// TIA Portal V20 export
// export: Created 2026-10-19T18:42:36.9079896Z, ExportSetting WithDefaults, DisplayName Totally Integrated Automation Portal, DisplayVersion V20 Update 6, DisplayName TIA Portal Openness, DisplayVersion V20 Update 6, DisplayName TIA Portal Version Control Interface, DisplayVersion V20 Update 6, DisplayName SINAMICS Startdrive Advanced, DisplayVersion V20 SP1, DisplayName SINAMICS Startdrive G130, G150, S120, S150, SINAMICS MV, G220, S200, S210, DisplayVersion V20 SP1, DisplayName SINAMICS Startdrive G110M, G120, G120C, G120D, G120P, G115D, DisplayVersion V20 SP1, DisplayName STEP 7 Professional, DisplayVersion V20 Update 6, DisplayName STEP 7 Safety, DisplayVersion V20 Update 2, DisplayName WinCC Basic/Comfort/Advanced, DisplayVersion V20 Update 6, DisplayName WinCC Unified, DisplayVersion V20 Update 6
FUNCTION_BLOCK "Remote_Panel"   // FB17, F_LAD
{ S7_Optimized_Access := 'TRUE' }
VERSION : 0.1
// stored: AutoNumber true, IsIECCheckEnabled false, UDAEnableTagReadback false
   VAR_INPUT
      ID : Int;
      Overtravel_Lower_limit : Bool;
      Overtravel_Upper_limit : Bool;
      Estop : Bool;
      Reset : Bool;
      Chain_Slack_1 : Bool;
      Chain_Slack_2 : Bool;
      Chain_Slack_3 : Bool;
      Chain_Slack_4 : Bool;
      "Light Guards 1" : Bool;
      "Light Guards 2" : Bool;
      Gate_1 : Bool;
      Gate_2 : Bool;
      EStop_Lock_1 : Bool;
      EStop_Lock_2 : Bool;
      Lock_Secured_1 : Bool;
      Lock_Secured_2 : Bool;
      "EStop Level 1" : Bool;
      "EStop Level 2" : Bool;
      "EStop Level 3" : Bool;
      "EStop Level 4" : Bool;
      "EStop Level 5" : Bool;
      "EStop Level 6" : Bool;
      Bypass : "F_Bypass_RemotePanel";
   END_VAR
   VAR_OUTPUT
      Safety_OK : Bool;
      Bypass_Warning : Bool;
      "STO VTD - CH1" : Bool;
      "STO VTD - CH2" : Bool;
      ACK { ExternalAccessible := 'False'; ExternalVisible := 'False'; ExternalWritable := 'False'} : Bool;
      L1_OK : Bool;
      L2_OK : Bool;
      L3_OK : Bool;
      L4_OK : Bool;
      L5_OK : Bool;
      L6_OK : Bool;
   END_VAR
   VAR
      Overtravel_Lower_Limit_DB : ESTOP1;
      Overtravel_Upper_Limit_DB : ESTOP1;
      Estop_Cabinet_DB : ESTOP1;
      Chain_Slack_1_DB : ESTOP1;
      Chain_Slack_2_DB : ESTOP1;
      Chain_Slack_3_DB : ESTOP1;
      Chain_Slack_4_DB : ESTOP1;
      "Light_Guards 1" : ESTOP1;
      "Light_Guards 2" : ESTOP1;
      Gate_1_DB : ESTOP1;
      Gate_2_DB : ESTOP1;
      EStop_Lock_1_DB : ESTOP1;
      EStop_Lock_2_DB : ESTOP1;
      Lock_Secured_1_DB : ESTOP1;
      Lock_Secured_2_DB : ESTOP1;
      "EStop Level 1_DB" : ESTOP1;
      "EStop Level 2_DB" : ESTOP1;
      "EStop Level 3_DB" : ESTOP1;
      "EStop Level 4_DB" : ESTOP1;
      "EStop Level 5_DB" : ESTOP1;
      "EStop Level 6_DB" : ESTOP1;
   END_VAR
   VAR_TEMP
      EStop_Levels_OK : Bool;
   END_VAR
BEGIN

REGION Network 1: RESET CABINET
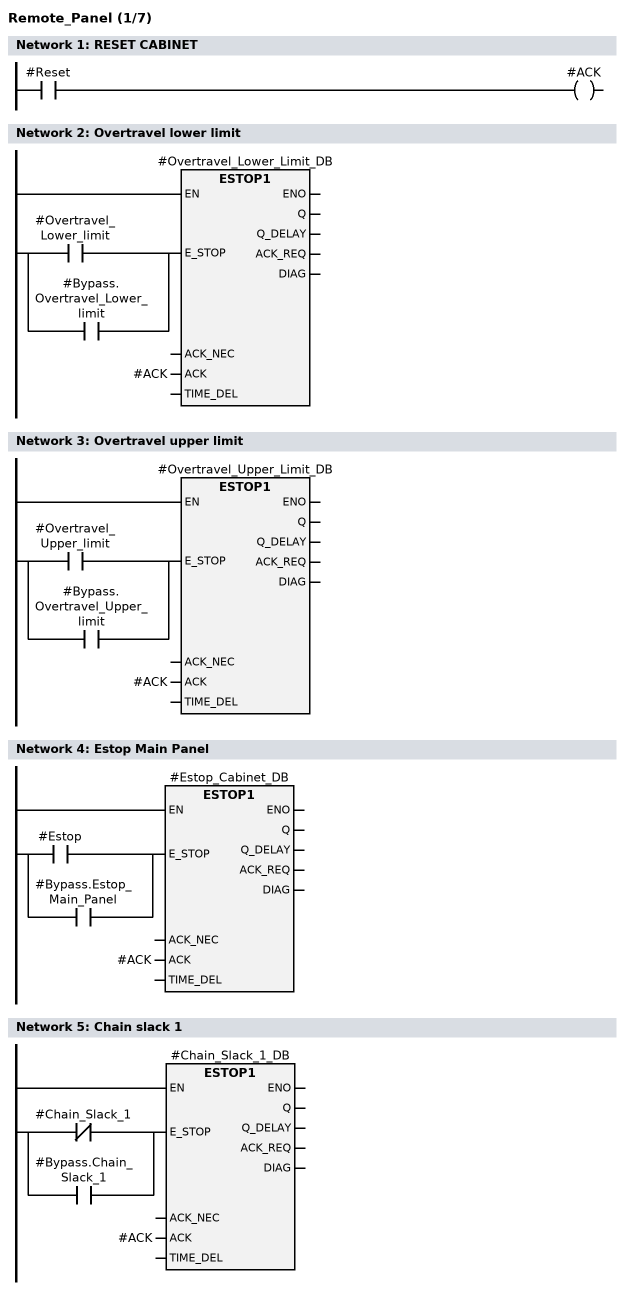
   RUNG wire#powerrail
      Contact( #Reset )
      Coil( #ACK )
   END_RUNG
   // the same network as SCL:
   #ACK := #Reset;
END_REGION

REGION Network 2: Overtravel lower limit
   RUNG wire#powerrail
      #Overtravel_Lower_Limit_DB.ESTOP1(E_STOP := wire#w1, ACK_NEC :=, ACK := #ACK, TIME_DEL :=, Q =>, Q_DELAY =>, ACK_REQ =>, DIAG =>)
   END_RUNG
   RUNG wire#powerrail
      Contact( #Overtravel_Lower_limit )
   END_RUNG wire#w1
   RUNG wire#powerrail
      Contact( #Bypass.Overtravel_Lower_limit )
   END_RUNG wire#w1
   // the same network as SCL:
   #Overtravel_Lower_Limit_DB(E_STOP := #Overtravel_Lower_limit OR #Bypass.Overtravel_Lower_limit, ACK := #ACK);   // ESTOP1
END_REGION

REGION Network 3: Overtravel upper limit
   RUNG wire#powerrail
      #Overtravel_Upper_Limit_DB.ESTOP1(E_STOP := wire#w1, ACK_NEC :=, ACK := #ACK, TIME_DEL :=, Q =>, Q_DELAY =>, ACK_REQ =>, DIAG =>)
   END_RUNG
   RUNG wire#powerrail
      Contact( #Overtravel_Upper_limit )
   END_RUNG wire#w1
   RUNG wire#powerrail
      Contact( #Bypass.Overtravel_Upper_limit )
   END_RUNG wire#w1
   // the same network as SCL:
   #Overtravel_Upper_Limit_DB(E_STOP := #Overtravel_Upper_limit OR #Bypass.Overtravel_Upper_limit, ACK := #ACK);   // ESTOP1
END_REGION

REGION Network 4: Estop Main Panel
   RUNG wire#powerrail
      #Estop_Cabinet_DB.ESTOP1(E_STOP := wire#w1, ACK_NEC :=, ACK := #ACK, TIME_DEL :=, Q =>, Q_DELAY =>, ACK_REQ =>, DIAG =>)
   END_RUNG
   RUNG wire#powerrail
      Contact( #Estop )
   END_RUNG wire#w1
   RUNG wire#powerrail
      Contact( #Bypass.Estop_Main_Panel )
   END_RUNG wire#w1
   // the same network as SCL:
   #Estop_Cabinet_DB(E_STOP := #Estop OR #Bypass.Estop_Main_Panel, ACK := #ACK);   // ESTOP1
END_REGION

REGION Network 5: Chain slack 1
   RUNG wire#powerrail
      #Chain_Slack_1_DB.ESTOP1(E_STOP := wire#w1, ACK_NEC :=, ACK := #ACK, TIME_DEL :=, Q =>, Q_DELAY =>, ACK_REQ =>, DIAG =>)
   END_RUNG
   RUNG wire#powerrail
      I_Contact( #Chain_Slack_1 )
   END_RUNG wire#w1
   RUNG wire#powerrail
      Contact( #Bypass.Chain_Slack_1 )
   END_RUNG wire#w1
   // the same network as SCL:
   #Chain_Slack_1_DB(E_STOP := NOT #Chain_Slack_1 OR #Bypass.Chain_Slack_1, ACK := #ACK);   // ESTOP1
END_REGION

REGION Network 6: Chain slack 2
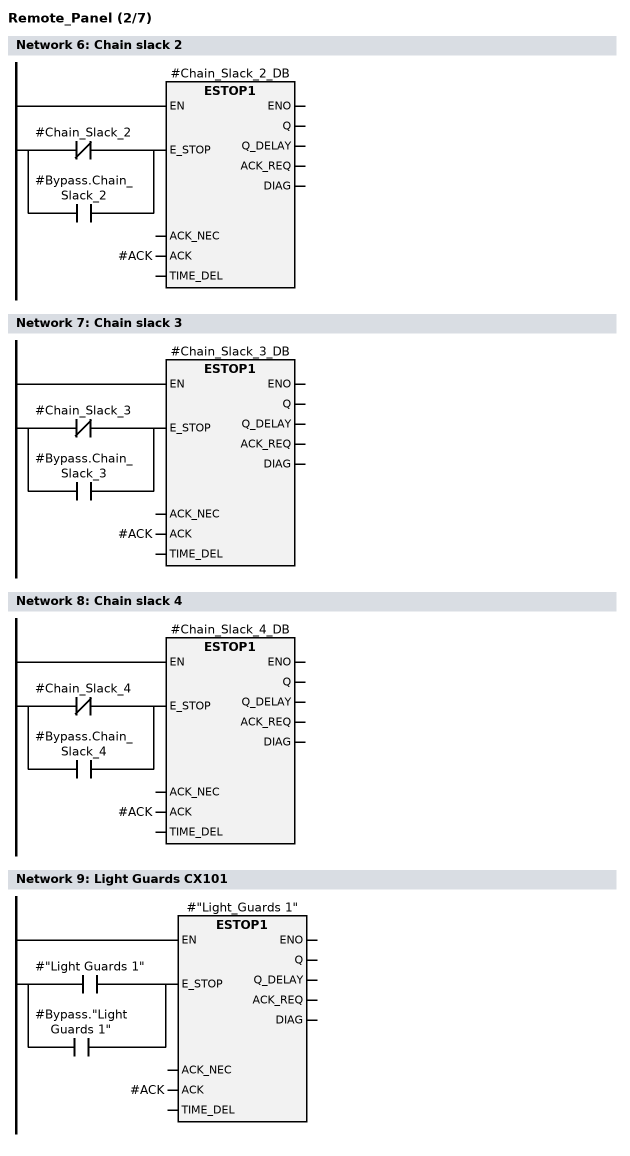
   RUNG wire#powerrail
      #Chain_Slack_2_DB.ESTOP1(E_STOP := wire#w1, ACK_NEC :=, ACK := #ACK, TIME_DEL :=, Q =>, Q_DELAY =>, ACK_REQ =>, DIAG =>)
   END_RUNG
   RUNG wire#powerrail
      I_Contact( #Chain_Slack_2 )
   END_RUNG wire#w1
   RUNG wire#powerrail
      Contact( #Bypass.Chain_Slack_2 )
   END_RUNG wire#w1
   // the same network as SCL:
   #Chain_Slack_2_DB(E_STOP := NOT #Chain_Slack_2 OR #Bypass.Chain_Slack_2, ACK := #ACK);   // ESTOP1
END_REGION

REGION Network 7: Chain slack 3
   RUNG wire#powerrail
      #Chain_Slack_3_DB.ESTOP1(E_STOP := wire#w1, ACK_NEC :=, ACK := #ACK, TIME_DEL :=, Q =>, Q_DELAY =>, ACK_REQ =>, DIAG =>)
   END_RUNG
   RUNG wire#powerrail
      I_Contact( #Chain_Slack_3 )
   END_RUNG wire#w1
   RUNG wire#powerrail
      Contact( #Bypass.Chain_Slack_3 )
   END_RUNG wire#w1
   // the same network as SCL:
   #Chain_Slack_3_DB(E_STOP := NOT #Chain_Slack_3 OR #Bypass.Chain_Slack_3, ACK := #ACK);   // ESTOP1
END_REGION

REGION Network 8: Chain slack 4
   RUNG wire#powerrail
      #Chain_Slack_4_DB.ESTOP1(E_STOP := wire#w1, ACK_NEC :=, ACK := #ACK, TIME_DEL :=, Q =>, Q_DELAY =>, ACK_REQ =>, DIAG =>)
   END_RUNG
   RUNG wire#powerrail
      I_Contact( #Chain_Slack_4 )
   END_RUNG wire#w1
   RUNG wire#powerrail
      Contact( #Bypass.Chain_Slack_4 )
   END_RUNG wire#w1
   // the same network as SCL:
   #Chain_Slack_4_DB(E_STOP := NOT #Chain_Slack_4 OR #Bypass.Chain_Slack_4, ACK := #ACK);   // ESTOP1
END_REGION

REGION Network 9: Light Guards CX101
   RUNG wire#powerrail
      #"Light_Guards 1".ESTOP1(E_STOP := wire#w1, ACK_NEC :=, ACK := #ACK, TIME_DEL :=, Q =>, Q_DELAY =>, ACK_REQ =>, DIAG =>)
   END_RUNG
   RUNG wire#powerrail
      Contact( #"Light Guards 1" )
   END_RUNG wire#w1
   RUNG wire#powerrail
      Contact( #Bypass."Light Guards 1" )
   END_RUNG wire#w1
   // the same network as SCL:
   #"Light_Guards 1"(E_STOP := #"Light Guards 1" OR #Bypass."Light Guards 1", ACK := #ACK);   // ESTOP1
END_REGION

REGION Network 10: Light Guards CX201
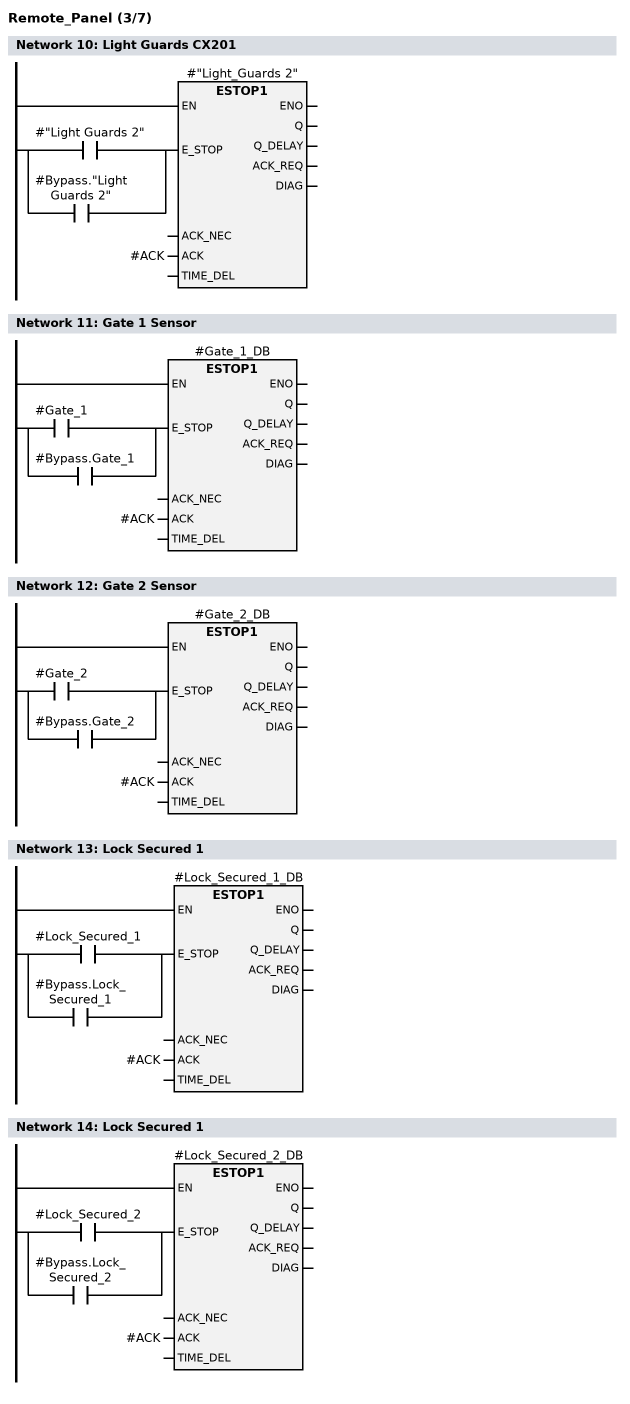
   RUNG wire#powerrail
      #"Light_Guards 2".ESTOP1(E_STOP := wire#w1, ACK_NEC :=, ACK := #ACK, TIME_DEL :=, Q =>, Q_DELAY =>, ACK_REQ =>, DIAG =>)
   END_RUNG
   RUNG wire#powerrail
      Contact( #"Light Guards 2" )
   END_RUNG wire#w1
   RUNG wire#powerrail
      Contact( #Bypass."Light Guards 2" )
   END_RUNG wire#w1
   // the same network as SCL:
   #"Light_Guards 2"(E_STOP := #"Light Guards 2" OR #Bypass."Light Guards 2", ACK := #ACK);   // ESTOP1
END_REGION

REGION Network 11: Gate 1 Sensor
   RUNG wire#powerrail
      #Gate_1_DB.ESTOP1(E_STOP := wire#w1, ACK_NEC :=, ACK := #ACK, TIME_DEL :=, Q =>, Q_DELAY =>, ACK_REQ =>, DIAG =>)
   END_RUNG
   RUNG wire#powerrail
      Contact( #Gate_1 )
   END_RUNG wire#w1
   RUNG wire#powerrail
      Contact( #Bypass.Gate_1 )
   END_RUNG wire#w1
   // the same network as SCL:
   #Gate_1_DB(E_STOP := #Gate_1 OR #Bypass.Gate_1, ACK := #ACK);   // ESTOP1
END_REGION

REGION Network 12: Gate 2 Sensor
   RUNG wire#powerrail
      #Gate_2_DB.ESTOP1(E_STOP := wire#w1, ACK_NEC :=, ACK := #ACK, TIME_DEL :=, Q =>, Q_DELAY =>, ACK_REQ =>, DIAG =>)
   END_RUNG
   RUNG wire#powerrail
      Contact( #Gate_2 )
   END_RUNG wire#w1
   RUNG wire#powerrail
      Contact( #Bypass.Gate_2 )
   END_RUNG wire#w1
   // the same network as SCL:
   #Gate_2_DB(E_STOP := #Gate_2 OR #Bypass.Gate_2, ACK := #ACK);   // ESTOP1
END_REGION

REGION Network 13: Lock Secured 1
   RUNG wire#powerrail
      #Lock_Secured_1_DB.ESTOP1(E_STOP := wire#w1, ACK_NEC :=, ACK := #ACK, TIME_DEL :=, Q =>, Q_DELAY =>, ACK_REQ =>, DIAG =>)
   END_RUNG
   RUNG wire#powerrail
      Contact( #Lock_Secured_1 )
   END_RUNG wire#w1
   RUNG wire#powerrail
      Contact( #Bypass.Lock_Secured_1 )
   END_RUNG wire#w1
   // the same network as SCL:
   #Lock_Secured_1_DB(E_STOP := #Lock_Secured_1 OR #Bypass.Lock_Secured_1, ACK := #ACK);   // ESTOP1
END_REGION

REGION Network 14: Lock Secured 1
   RUNG wire#powerrail
      #Lock_Secured_2_DB.ESTOP1(E_STOP := wire#w1, ACK_NEC :=, ACK := #ACK, TIME_DEL :=, Q =>, Q_DELAY =>, ACK_REQ =>, DIAG =>)
   END_RUNG
   RUNG wire#powerrail
      Contact( #Lock_Secured_2 )
   END_RUNG wire#w1
   RUNG wire#powerrail
      Contact( #Bypass.Lock_Secured_2 )
   END_RUNG wire#w1
   // the same network as SCL:
   #Lock_Secured_2_DB(E_STOP := #Lock_Secured_2 OR #Bypass.Lock_Secured_2, ACK := #ACK);   // ESTOP1
END_REGION

REGION Network 15: Idem Lock EStop 1
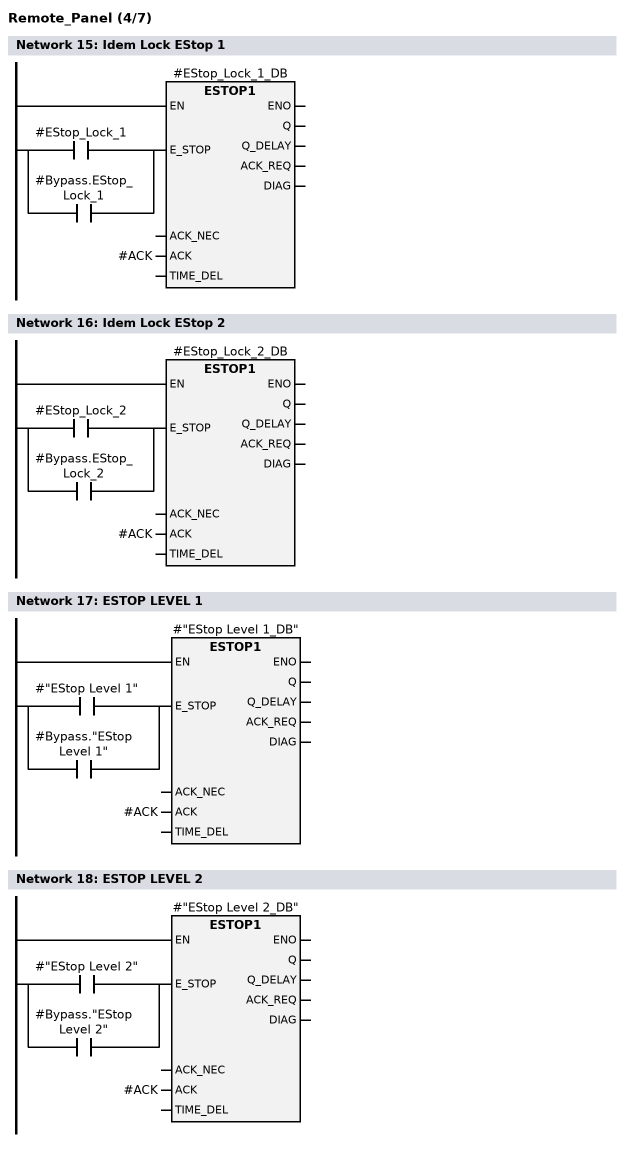
   RUNG wire#powerrail
      #EStop_Lock_1_DB.ESTOP1(E_STOP := wire#w1, ACK_NEC :=, ACK := #ACK, TIME_DEL :=, Q =>, Q_DELAY =>, ACK_REQ =>, DIAG =>)
   END_RUNG
   RUNG wire#powerrail
      Contact( #EStop_Lock_1 )
   END_RUNG wire#w1
   RUNG wire#powerrail
      Contact( #Bypass.EStop_Lock_1 )
   END_RUNG wire#w1
   // the same network as SCL:
   #EStop_Lock_1_DB(E_STOP := #EStop_Lock_1 OR #Bypass.EStop_Lock_1, ACK := #ACK);   // ESTOP1
END_REGION

REGION Network 16: Idem Lock EStop 2
   RUNG wire#powerrail
      #EStop_Lock_2_DB.ESTOP1(E_STOP := wire#w1, ACK_NEC :=, ACK := #ACK, TIME_DEL :=, Q =>, Q_DELAY =>, ACK_REQ =>, DIAG =>)
   END_RUNG
   RUNG wire#powerrail
      Contact( #EStop_Lock_2 )
   END_RUNG wire#w1
   RUNG wire#powerrail
      Contact( #Bypass.EStop_Lock_2 )
   END_RUNG wire#w1
   // the same network as SCL:
   #EStop_Lock_2_DB(E_STOP := #EStop_Lock_2 OR #Bypass.EStop_Lock_2, ACK := #ACK);   // ESTOP1
END_REGION

REGION Network 17: ESTOP LEVEL 1
   RUNG wire#powerrail
      #"EStop Level 1_DB".ESTOP1(E_STOP := wire#w1, ACK_NEC :=, ACK := #ACK, TIME_DEL :=, Q =>, Q_DELAY =>, ACK_REQ =>, DIAG =>)
   END_RUNG
   RUNG wire#powerrail
      Contact( #"EStop Level 1" )
   END_RUNG wire#w1
   RUNG wire#powerrail
      Contact( #Bypass."EStop Level 1" )
   END_RUNG wire#w1
   // the same network as SCL:
   #"EStop Level 1_DB"(E_STOP := #"EStop Level 1" OR #Bypass."EStop Level 1", ACK := #ACK);   // ESTOP1
END_REGION

REGION Network 18: ESTOP LEVEL 2
   RUNG wire#powerrail
      #"EStop Level 2_DB".ESTOP1(E_STOP := wire#w1, ACK_NEC :=, ACK := #ACK, TIME_DEL :=, Q =>, Q_DELAY =>, ACK_REQ =>, DIAG =>)
   END_RUNG
   RUNG wire#powerrail
      Contact( #"EStop Level 2" )
   END_RUNG wire#w1
   RUNG wire#powerrail
      Contact( #Bypass."EStop Level 2" )
   END_RUNG wire#w1
   // the same network as SCL:
   #"EStop Level 2_DB"(E_STOP := #"EStop Level 2" OR #Bypass."EStop Level 2", ACK := #ACK);   // ESTOP1
END_REGION

REGION Network 19: ESTOP LEVEL 3
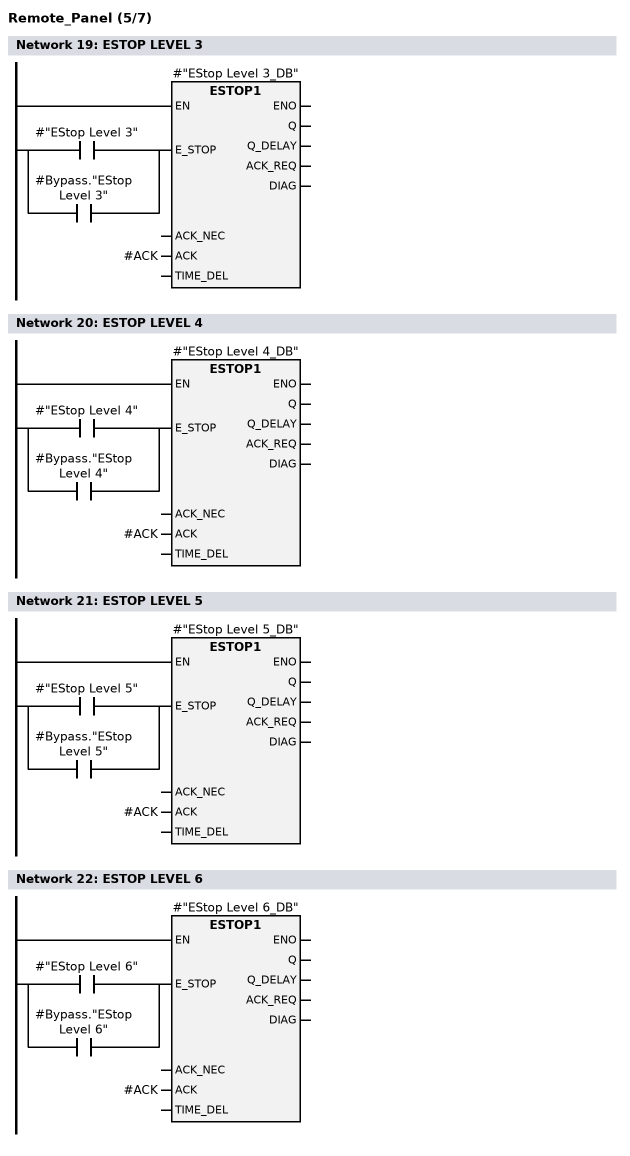
   RUNG wire#powerrail
      #"EStop Level 3_DB".ESTOP1(E_STOP := wire#w1, ACK_NEC :=, ACK := #ACK, TIME_DEL :=, Q =>, Q_DELAY =>, ACK_REQ =>, DIAG =>)
   END_RUNG
   RUNG wire#powerrail
      Contact( #"EStop Level 3" )
   END_RUNG wire#w1
   RUNG wire#powerrail
      Contact( #Bypass."EStop Level 3" )
   END_RUNG wire#w1
   // the same network as SCL:
   #"EStop Level 3_DB"(E_STOP := #"EStop Level 3" OR #Bypass."EStop Level 3", ACK := #ACK);   // ESTOP1
END_REGION

REGION Network 20: ESTOP LEVEL 4
   RUNG wire#powerrail
      #"EStop Level 4_DB".ESTOP1(E_STOP := wire#w1, ACK_NEC :=, ACK := #ACK, TIME_DEL :=, Q =>, Q_DELAY =>, ACK_REQ =>, DIAG =>)
   END_RUNG
   RUNG wire#powerrail
      Contact( #"EStop Level 4" )
   END_RUNG wire#w1
   RUNG wire#powerrail
      Contact( #Bypass."EStop Level 4" )
   END_RUNG wire#w1
   // the same network as SCL:
   #"EStop Level 4_DB"(E_STOP := #"EStop Level 4" OR #Bypass."EStop Level 4", ACK := #ACK);   // ESTOP1
END_REGION

REGION Network 21: ESTOP LEVEL 5
   RUNG wire#powerrail
      #"EStop Level 5_DB".ESTOP1(E_STOP := wire#w1, ACK_NEC :=, ACK := #ACK, TIME_DEL :=, Q =>, Q_DELAY =>, ACK_REQ =>, DIAG =>)
   END_RUNG
   RUNG wire#powerrail
      Contact( #"EStop Level 5" )
   END_RUNG wire#w1
   RUNG wire#powerrail
      Contact( #Bypass."EStop Level 5" )
   END_RUNG wire#w1
   // the same network as SCL:
   #"EStop Level 5_DB"(E_STOP := #"EStop Level 5" OR #Bypass."EStop Level 5", ACK := #ACK);   // ESTOP1
END_REGION

REGION Network 22: ESTOP LEVEL 6
   RUNG wire#powerrail
      #"EStop Level 6_DB".ESTOP1(E_STOP := wire#w1, ACK_NEC :=, ACK := #ACK, TIME_DEL :=, Q =>, Q_DELAY =>, ACK_REQ =>, DIAG =>)
   END_RUNG
   RUNG wire#powerrail
      Contact( #"EStop Level 6" )
   END_RUNG wire#w1
   RUNG wire#powerrail
      Contact( #Bypass."EStop Level 6" )
   END_RUNG wire#w1
   // the same network as SCL:
   #"EStop Level 6_DB"(E_STOP := #"EStop Level 6" OR #Bypass."EStop Level 6", ACK := #ACK);   // ESTOP1
END_REGION

REGION Network 23: STOP LEVEL
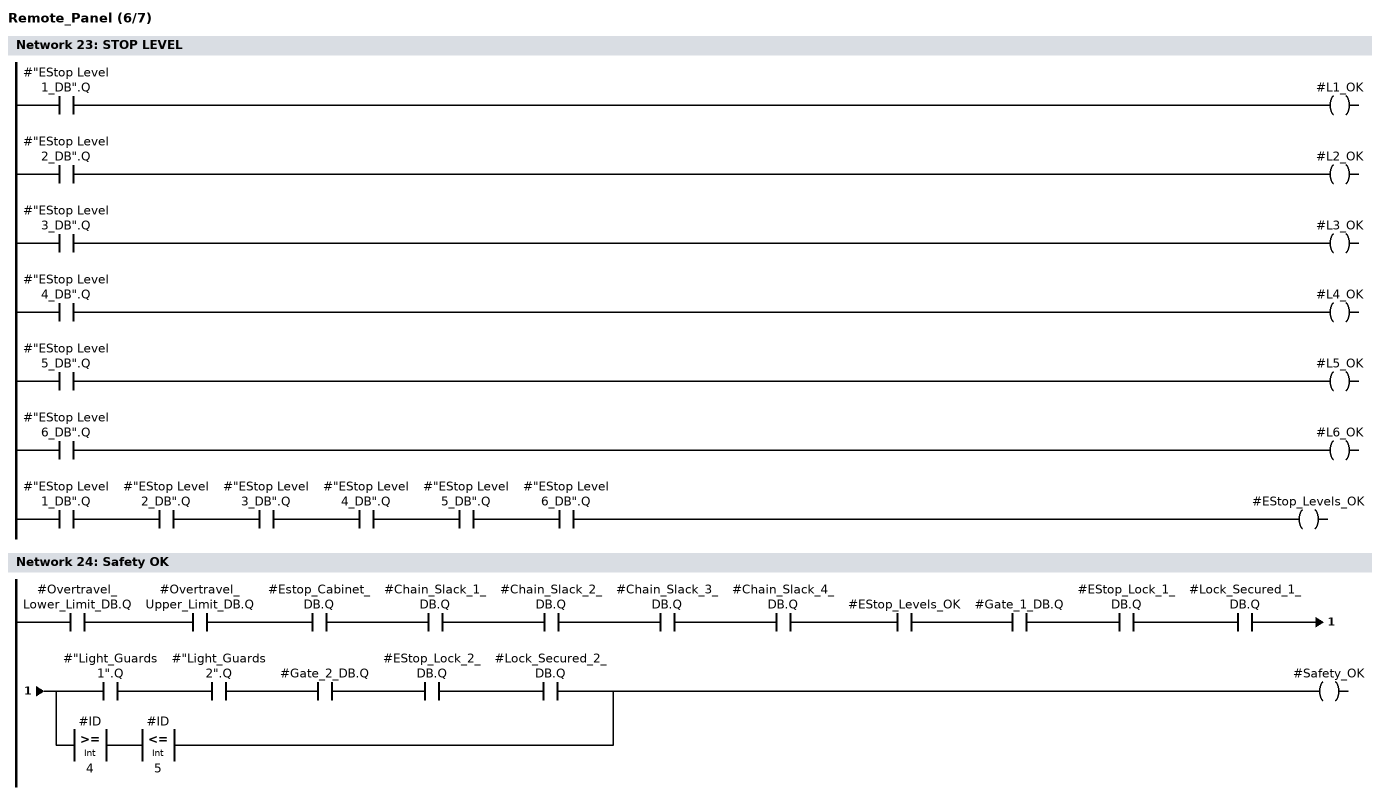
   RUNG wire#powerrail
      Contact( #"EStop Level 1_DB".Q )
      Coil( #L1_OK )
   END_RUNG
   RUNG wire#powerrail
      Contact( #"EStop Level 2_DB".Q )
      Coil( #L2_OK )
   END_RUNG
   RUNG wire#powerrail
      Contact( #"EStop Level 3_DB".Q )
      Coil( #L3_OK )
   END_RUNG
   RUNG wire#powerrail
      Contact( #"EStop Level 4_DB".Q )
      Coil( #L4_OK )
   END_RUNG
   RUNG wire#powerrail
      Contact( #"EStop Level 5_DB".Q )
      Coil( #L5_OK )
   END_RUNG
   RUNG wire#powerrail
      Contact( #"EStop Level 6_DB".Q )
      Coil( #L6_OK )
   END_RUNG
   RUNG wire#powerrail
      Contact( #"EStop Level 1_DB".Q )
      Contact( #"EStop Level 2_DB".Q )
      Contact( #"EStop Level 3_DB".Q )
      Contact( #"EStop Level 4_DB".Q )
      Contact( #"EStop Level 5_DB".Q )
      Contact( #"EStop Level 6_DB".Q )
      Coil( #EStop_Levels_OK )
   END_RUNG
   // the same network as SCL:
   #L1_OK := #"EStop Level 1_DB".Q;
   #L2_OK := #"EStop Level 2_DB".Q;
   #L3_OK := #"EStop Level 3_DB".Q;
   #L4_OK := #"EStop Level 4_DB".Q;
   #L5_OK := #"EStop Level 5_DB".Q;
   #L6_OK := #"EStop Level 6_DB".Q;
   #EStop_Levels_OK := #"EStop Level 1_DB".Q AND #"EStop Level 2_DB".Q AND #"EStop Level 3_DB".Q AND #"EStop Level 4_DB".Q AND #"EStop Level 5_DB".Q AND #"EStop Level 6_DB".Q;
END_REGION

REGION Network 24: Safety OK
   RUNG wire#powerrail
      Contact( #Overtravel_Lower_Limit_DB.Q )
      Contact( #Overtravel_Upper_Limit_DB.Q )
      Contact( #Estop_Cabinet_DB.Q )
      Contact( #Chain_Slack_1_DB.Q )
      Contact( #Chain_Slack_2_DB.Q )
      Contact( #Chain_Slack_3_DB.Q )
      Contact( #Chain_Slack_4_DB.Q )
      Contact( #EStop_Levels_OK )
      Contact( #Gate_1_DB.Q )
      Contact( #EStop_Lock_1_DB.Q )
      Contact( #Lock_Secured_1_DB.Q )
      wire#w1
      Contact( #"Light_Guards 1".Q )
      Contact( #"Light_Guards 2".Q )
      Contact( #Gate_2_DB.Q )
      Contact( #EStop_Lock_2_DB.Q )
      Contact( #Lock_Secured_2_DB.Q )
      wire#w2
      Coil( #Safety_OK )
   END_RUNG
   RUNG wire#w1
      { S7_Templates := "SrcType := Int" } GE_Contact(in1 := #ID, in2 := 4)
      { S7_Templates := "SrcType := Int" } LE_Contact(in1 := #ID, in2 := 5)
   END_RUNG wire#w2
   // the same network as SCL:
   #Safety_OK := #Overtravel_Lower_Limit_DB.Q AND #Overtravel_Upper_Limit_DB.Q AND #Estop_Cabinet_DB.Q AND #Chain_Slack_1_DB.Q AND #Chain_Slack_2_DB.Q AND #Chain_Slack_3_DB.Q AND #Chain_Slack_4_DB.Q AND #EStop_Levels_OK AND #Gate_1_DB.Q AND #EStop_Lock_1_DB.Q AND #Lock_Secured_1_DB.Q AND ((#"Light_Guards 1".Q AND #"Light_Guards 2".Q AND #Gate_2_DB.Q AND #EStop_Lock_2_DB.Q AND #Lock_Secured_2_DB.Q) OR ((#ID >= 4) AND (#ID <= 5)));
END_REGION

REGION Network 25: Bypass Warning
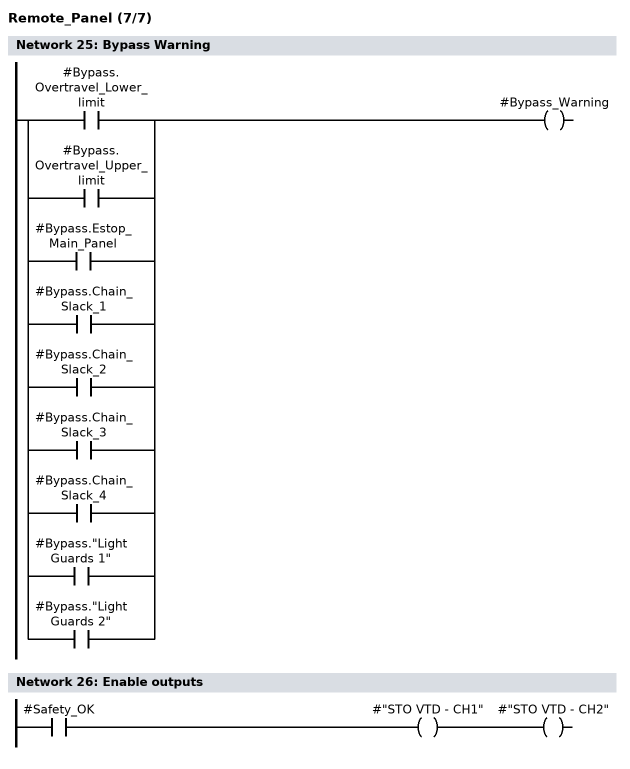
   RUNG wire#powerrail
      Contact( #Bypass.Overtravel_Lower_limit )
      wire#w1
      Coil( #Bypass_Warning )
   END_RUNG
   RUNG wire#powerrail
      Contact( #Bypass.Overtravel_Upper_limit )
   END_RUNG wire#w1
   RUNG wire#powerrail
      Contact( #Bypass.Estop_Main_Panel )
   END_RUNG wire#w1
   RUNG wire#powerrail
      Contact( #Bypass.Chain_Slack_1 )
   END_RUNG wire#w1
   RUNG wire#powerrail
      Contact( #Bypass.Chain_Slack_2 )
   END_RUNG wire#w1
   RUNG wire#powerrail
      Contact( #Bypass.Chain_Slack_3 )
   END_RUNG wire#w1
   RUNG wire#powerrail
      Contact( #Bypass.Chain_Slack_4 )
   END_RUNG wire#w1
   RUNG wire#powerrail
      Contact( #Bypass."Light Guards 1" )
   END_RUNG wire#w1
   RUNG wire#powerrail
      Contact( #Bypass."Light Guards 2" )
   END_RUNG wire#w1
   // the same network as SCL:
   #Bypass_Warning := #Bypass.Overtravel_Lower_limit OR #Bypass.Overtravel_Upper_limit OR #Bypass.Estop_Main_Panel OR #Bypass.Chain_Slack_1 OR #Bypass.Chain_Slack_2 OR #Bypass.Chain_Slack_3 OR #Bypass.Chain_Slack_4 OR #Bypass."Light Guards 1" OR #Bypass."Light Guards 2";
END_REGION

REGION Network 26: Enable outputs
   RUNG wire#powerrail
      Contact( #Safety_OK )
      Coil( #"STO VTD - CH1" )
      Coil( #"STO VTD - CH2" )
   END_RUNG
   // the same network as SCL:
   #"STO VTD - CH1" := #Safety_OK;
   #"STO VTD - CH2" := #Safety_OK;
END_REGION
END_FUNCTION_BLOCK
